// TIA Portal V21 export
// export: Created 2026-11-07T17:04:58.9997488Z, ExportSetting WithDefaults, DisplayName Totally Integrated Automation Portal, DisplayVersion V21, DisplayName STEP 7 Professional, DisplayVersion V21, DisplayName STEP 7 Safety, DisplayVersion V21, DisplayName Tech WebApplication, DisplayVersion V21, DisplayName WinCC Basic/Comfort/Advanced, DisplayVersion V21, DisplayName WinCC Unified, DisplayVersion V21
TextList "TL_Kind"  ListRange=Decimal
  TextListEntry   EntryType=SingleValue, Text="-"
  TextListEntry   EntryType=SingleValue, From=1, To=1, Text="ISTOVAR Bay0->Bay1"
  TextListEntry   EntryType=SingleValue, From=2, To=2, Text="UKRCAJ Bay1->Bay0"
